(*
SPDX-FileCopyrightText: © 2026 Oleksandr Tiutyk <trofimich@gmail.com>
SPDX-License-Identifier: MIT
License: https://opensource.org/license/mit
*)

(*!
<summary>Provides finite bounds for UnsignedByte values.</summary>
<description>
MIN_VALUE and MAX_VALUE describe the represented integer range; constants perform no conversion or runtime
validation. Additional named bounds, where declared, describe narrower representations.
</description>
*)

{attribute 'no_explicit_call' := 'do not call this function block directly'}
PROGRAM UnsignedInt8
VAR CONSTANT
	ZERO : USINT := 0;
	MIN_VALUE : USINT := 0;
	MAX_VALUE : USINT := BYTE#16#FF;
END_VAR
VAR
	{attribute 'hide'} 
	_ClassName : STRING := __POUNAME();
END_VAR

{attribute 'monitoring' := 'call'}
PROPERTY ClassName : REFERENCE TO STRING
GET
ClassName REF= _ClassName;
END_GET
END_PROPERTY

(*!
<summary>Provides the library namespace used in diagnostics.</summary>
<description>
Borrowed read-only reference to the compiler-initialized library namespace; no ownership transfer.
</description>
*)
{attribute 'monitoring' := 'call'}
PROPERTY NamespaceName : REFERENCE TO STRING
GET
NamespaceName REF= CurrentNamespace.Name;
END_GET
END_PROPERTY

END_PROGRAM

(* stored: Version 1.1.0.1
   POU UnsignedInt8: Id {4535912c-7c28-45af-ab90-74f12bea42b1}, SpecialFunc None
   Property ClassName: Id {7cdfd4b8-4143-436d-8a80-d8d11af812c3}
   Get Get: Id {a66bdd50-80ee-42c4-8efa-220958ec5c8a}
   Property NamespaceName: Id {7eb551b0-be22-4fd0-8050-6706a2730601}
   Get Get: Id {53ee3327-4ef7-469b-8356-c1c023ceb189} *)
